Fanuc KAREL source: KT00994.KL

PROGRAM KT00994
%NOLOCKGROUP
VAR
  P1: JOINTPOS
  P2: JOINTPOS
  X: REAL
  Y: REAL
  Z: REAL
  W: REAL
  P: REAL
  R: REAL
  CFG: CONFIG
BEGIN
  UNPOS(P1, X, Y, Z, W, P, R, CFG)
END KT00994
